TYPE ST_PolarIIChamber_HolderServiceStatus :
STRUCT
	Gripper : ST_PolarIIChamber_OpenCloseServiceStatus;
	Rotate : ST_PolarIIChamber_HolderRotateServiceStatus;
	VacuumEstablish : ST_ServiceStatus;
END_STRUCT
END_TYPE

(* stored: Version 1.1.0.1, ProductVersion 3.1.4026.18
   DUT ST_PolarIIChamber_HolderServiceStatus: Id {14000000-0000-0000-0000-000000000066} *)
